Fanuc KAREL source: KT00172.KL

PROGRAM KT00172
%NOLOCKGROUP
VAR
  R1: REAL
  R2: REAL
  OUT: REAL
BEGIN
  R1 = 2.0
  R2 = 3.0
  R1 = 2.0
  R2 = 3.0
  OUT = R1 MOD R2
END KT00172
